(* IEC 61131-3 sources: plcassist-cli/packages/volt-lsp-iec/test-corpus/pro2193/Device/Plc Logic/Application/09 Misc/Library Manager/L_USPP_SignalProcessing, 27 files *)

(* ---- GETBOOLEANPROPERTY.fun ---- *)
FUNCTION GETBOOLEANPROPERTY : BOOL
VAR_INPUT
	STKEY : WSTRING;
END_VAR
END_FUNCTION

(* ---- GETCOMPANY.fun ---- *)
FUNCTION GETCOMPANY : WSTRING
END_FUNCTION

(* ---- GETNUMBERPROPERTY.fun ---- *)
FUNCTION GETNUMBERPROPERTY : DINT
VAR_INPUT
	STKEY : WSTRING;
END_VAR
END_FUNCTION

(* ---- GETTEXTPROPERTY.fun ---- *)
FUNCTION GETTEXTPROPERTY : WSTRING
VAR_INPUT
	STKEY : WSTRING;
END_VAR
END_FUNCTION

(* ---- GETTEXTPROPERTY2.fun ---- *)
FUNCTION GETTEXTPROPERTY2 : POINTER TO WSTRING
VAR_INPUT
	STKEY : WSTRING;
END_VAR
END_FUNCTION

(* ---- GETTITLE.fun ---- *)
FUNCTION GETTITLE : WSTRING
END_FUNCTION

(* ---- GETVERSION.fun ---- *)
FUNCTION GETVERSION : VERSION
END_FUNCTION

(* ---- GETVERSIONPROPERTY.fun ---- *)
FUNCTION GETVERSIONPROPERTY : VERSION
VAR_INPUT
	STKEY : WSTRING;
END_VAR
END_FUNCTION

(* ---- L_USPP_HLPPT1FILT.fun ---- *)
FUNCTION L_USPP_HLPPT1FILT : LREAL
VAR_INPUT
	LRVALUE : LREAL;
	LRINPUT : LREAL;
	LRNEW_N : LREAL;
END_VAR
END_FUNCTION

(* ---- GLOBALTEXTLIST.fb ---- *)
FUNCTION_BLOCK GLOBALTEXTLIST
VAR
	M_TEXTLISTFILE : STRING(255);
	_STNAMESPACE : STRING;
END_VAR
END_FUNCTION_BLOCK

(* ---- IMAGEPOOL.fb ---- *)
FUNCTION_BLOCK IMAGEPOOL
VAR
	M_STNAMESPACE : STRING(80);
	M_STHELPVARID : STRING;
	M_STHELPVARPATH : STRING(255);
	M_STHELP : STRING;
	M_REGISTERIMAGES : BOOL := TRUE;
END_VAR
END_FUNCTION_BLOCK

METHOD FB_INIT : BOOL
VAR_INPUT
	BINITRETAINS : BOOL;
	BINCOPYCODE : BOOL;
END_VAR
END_METHOD

METHOD FB_REINIT : BOOL
END_METHOD

METHOD FB_EXIT : BOOL
VAR_INPUT
	BINCOPYCODE : BOOL;
END_VAR
END_METHOD

(* ---- L_USPP_AVERAGEFILTER.fb ---- *)
FUNCTION_BLOCK L_USPP_AVERAGEFILTER EXTENDS L_USPP_Filter
VAR_INPUT
	LRFILTERTIME : LREAL;
	XCALCFILTERDELAY : BOOL := TRUE;
END_VAR
VAR_OUTPUT
	LRFILTERDELAY : LREAL;
END_VAR
VAR
	_ITFMEMORY : L_UBUP_IMemoryProvider;
	_DWDIM : DWORD;
	_DWBUFFERCOUNT : DWORD;
	_DWACTFILTERDEPTH : DWORD;
	_DWBUFFERSIZE : DWORD;
	_DWMEMSIZE : DWORD;
	_DWACTBUFFERPOS : DWORD;
	_DWPREVBUFFERPOS : DWORD;
	_DWVALIDDATA : DWORD;
	_ALRPTRBUFFER : ARRAY [0..(dwMaxDeriv + 1)] OF POINTER TO LREAL;
	_ONE_OVER_N : LREAL;
	_XFIRSTROUNDDONE : BOOL;
	_DWSTANDSTILLCNT : DWORD;
	_ALRFILTERED : ARRAY [0..dwMaxDeriv] OF LREAL;
END_VAR
END_FUNCTION_BLOCK

METHOD CYCLICACTION
VAR_INPUT
	ITFTIMINGCONTROLLER : L_UBUP.L_UBUP_ITimingController;
END_VAR
VAR_OUTPUT
	XCOMPLETE : BOOL;
	XABORT : BOOL;
	IERRORID : INT;
END_VAR
END_METHOD

METHOD RESETACTION
VAR_OUTPUT
	XCOMPLETE : BOOL;
END_VAR
END_METHOD

METHOD STARTACTION
VAR_OUTPUT
	XCOMPLETE : BOOL;
	IERRORID : INT;
END_VAR
END_METHOD

METHOD EVALMEMORYPROVIDER
VAR_INPUT
	ITFMEMORYPROVIDER : L_UBUP_IMemoryProvider;
END_VAR
END_METHOD

METHOD FB_INIT : BOOL
VAR_INPUT
	BINITRETAINS : BOOL;
	BINCOPYCODE : BOOL;
	DWDERIVS : DWORD;
	ITFMEMORY : L_UBUP_IMemoryProvider;
END_VAR
END_METHOD

METHOD FILTERDELAY : LREAL
VAR_INPUT
	LRROUNDS : LREAL;
	LRCYCLELENGTH : LREAL;
END_VAR
END_METHOD

METHOD DISTRIBUTEBUFFER
END_METHOD

METHOD FILTER
VAR_INPUT
	PLR : POINTER TO LREAL;
END_VAR
VAR_IN_OUT
	LRFILTERED : LREAL;
END_VAR
END_METHOD

METHOD FILTERDETECTOVERFLOW
VAR_INPUT
	LRNEXTPOS : LREAL;
	LRPREVPOS : LREAL;
	LRMODCYCLE : LREAL;
END_VAR
VAR_OUTPUT
	LRMODCYCLENEW : LREAL;
END_VAR
END_METHOD

METHOD FILTERMODULO
END_METHOD

METHOD FILTEROUTPUT
VAR_IN_OUT
	ALRFILTERED : ARRAY [0..dwMaxDeriv] OF LREAL;
	ALROUTPUT : ARRAY [0..dwMaxDeriv] OF LREAL;
END_VAR
END_METHOD

(* ---- L_USPP_AVERAGEFILTEREXPLICIT.fb ---- *)
FUNCTION_BLOCK L_USPP_AVERAGEFILTEREXPLICIT EXTENDS L_USPP_AverageFilter
END_FUNCTION_BLOCK

METHOD FB_INIT : BOOL
VAR_INPUT
	BINITRETAINS : BOOL;
	BINCOPYCODE : BOOL;
	DWDERIVS : DWORD;
	ITFMEMORY : L_UBUP_IMemoryProvider;
END_VAR
END_METHOD

METHOD FILTER
VAR_INPUT
	PLR : POINTER TO LREAL;
END_VAR
VAR_IN_OUT
	LRFILTERED : LREAL;
END_VAR
END_METHOD

METHOD FILTERMODULO
END_METHOD

(* ---- L_USPP_AVERAGEFILTERRECURSIVE.fb ---- *)
FUNCTION_BLOCK L_USPP_AVERAGEFILTERRECURSIVE EXTENDS L_USPP_AverageFilter
VAR
	_XALLOWMODULO : BOOL;
END_VAR
END_FUNCTION_BLOCK

METHOD STARTACTION
VAR_OUTPUT
	XCOMPLETE : BOOL;
	IERRORID : INT;
END_VAR
END_METHOD

METHOD FB_INIT : BOOL
VAR_INPUT
	BINITRETAINS : BOOL;
	BINCOPYCODE : BOOL;
	DWDERIVS : DWORD;
	ITFMEMORY : L_UBUP_IMemoryProvider;
	XALLOWMODULO : BOOL;
END_VAR
END_METHOD

METHOD FILTERROUNDSCOUNTING
END_METHOD

METHOD FILTER
VAR_INPUT
	PLR : POINTER TO LREAL;
END_VAR
VAR_IN_OUT
	LRFILTERED : LREAL;
END_VAR
END_METHOD

METHOD FILTERMODULO
END_METHOD

METHOD FILTEROUTPUT
VAR_IN_OUT
	ALRFILTERED : ARRAY [0..dwMaxDeriv] OF LREAL;
	ALROUTPUT : ARRAY [0..dwMaxDeriv] OF LREAL;
END_VAR
END_METHOD

(* ---- L_USPP_BUTTERWORTH2NDORDER.fb ---- *)
FUNCTION_BLOCK L_USPP_BUTTERWORTH2NDORDER
VAR_INPUT
	LRIN : LREAL;
	LRFILTERTIME : LREAL;
	LRSAMPLINGTIME : LREAL;
	XINITWITHFIRSTINPUTVALUE : BOOL;
END_VAR
VAR_OUTPUT
	LROUT : LREAL;
END_VAR
VAR
	_LRINITCYCLETIME : LREAL;
	_LRFILTERTIME : LREAL;
	LRTASKCYCLE : LREAL;
	LROMEGA : LREAL;
	ALRXINT : ARRAY [0..2] OF LREAL;
	ALRYINT : ARRAY [0..2] OF LREAL;
	LRB0 : LREAL;
	LRB1 : LREAL;
	LRB2 : LREAL;
	LRA0 : LREAL;
	LRA0INV : LREAL;
	LRA1 : LREAL;
	LRA2 : LREAL;
	LROMEGASQUARED : LREAL;
	C_LRSQRT2 : LREAL := SQRT(2);
END_VAR
END_FUNCTION_BLOCK

METHOD FB_INIT : BOOL
VAR_INPUT
	BINITRETAINS : BOOL;
	BINCOPYCODE : BOOL;
END_VAR
END_METHOD

(* ---- L_USPP_COMPARE.fb ---- *)
FUNCTION_BLOCK L_USPP_COMPARE
VAR_INPUT
	LRIN1 : LREAL := 0;
	LRIN2 : LREAL := 0;
	DWFUNCTION : DWORD := 0;
	LRTOLERANCE : LREAL := 0;
	LRHYSTERESIS : LREAL := 0;
END_VAR
VAR_OUTPUT
	XOUT : BOOL := FALSE;
	XERROR : BOOL := FALSE;
	EERRORID : L_IE1P_Error;
END_VAR
VAR
	LRINTHYSTERESIS : LREAL := 0;
	LRINTWINDOW : LREAL := 0;
	LRINTIN1 : LREAL := 0;
	LRINTIN2 : LREAL := 0;
	LRINTTEMP : LREAL := 0;
	OUTVAR : BOOL;
END_VAR
END_FUNCTION_BLOCK

(* ---- L_USPP_CURVE.fb ---- *)
FUNCTION_BLOCK L_USPP_CURVE
VAR_INPUT
	LRIN : LREAL;
	DWMODE : DWORD;
	ALRXVALUES : ARRAY [1..9] OF LREAL;
	ALRYVALUES : ARRAY [1..9] OF LREAL;
END_VAR
VAR_OUTPUT
	LROUT : LREAL;
	XERROR : BOOL := FALSE;
	EERRORID : L_IE1P_Error;
END_VAR
VAR
	DISTARTIDX : DINT;
	DIENDIDX : DINT;
	LRLASTIN : LREAL;
	LRINPUT : LREAL;
	DISTART : DINT;
	DIEND : DINT;
	DITMP32 : DINT;
	XNEGINPUT : BOOL;
	XSAVELASTIN : BOOL;
	TMP : LREAL;
	GETMAXCURVEPOINTS : INT := 9;
END_VAR
END_FUNCTION_BLOCK

METHOD GETVALIDDATA
END_METHOD

(* ---- L_USPP_DEADTIMEINT.fb ---- *)
FUNCTION_BLOCK L_USPP_DEADTIMEINT
VAR_INPUT
	XENABLE : BOOL;
	XOFFSETACTIVE : BOOL;
	LRDELAY : LREAL;
	LRCYCLETIME : LREAL;
	PBIN : POINTER TO BYTE;
	PBOUT : POINTER TO BYTE;
	DISIZEOFDATA : DINT;
END_VAR
VAR_OUTPUT
	XBUSY : BOOL;
	XBUFFERINITIALIZED : BOOL;
	XERROR : BOOL;
	EERRORID : L_IE1P_Error;
END_VAR
VAR
	_XENABLEOLD : BOOL;
	_XOFFSETACTIVE : BOOL;
	_UDISIZEINT : UDINT;
	_LRCYCLETIME : LREAL;
	_LRINITCYCLETIME : LREAL;
	_WBUFFERCNT_1 : WORD;
	_WBUFFERCNT_2 : WORD;
	_WBUFFERLENGTH : WORD;
	_LRDELAY : LREAL;
	_LRRES : LREAL;
	_WDELAY : WORD;
	_PTMP : POINTER TO BYTE;
	_ITFMEMPROVIDER : L_UBUP_IMemoryProvider;
	_PBBUFFER : POINTER TO BYTE;
	_UDIBUFFERSIZE : UDINT;
END_VAR
END_FUNCTION_BLOCK

METHOD FB_INIT : BOOL
VAR_INPUT
	BINITRETAINS : BOOL;
	BINCOPYCODE : BOOL;
	ITFMEMPROVIDER : L_UBUP_IMemoryProvider;
END_VAR
END_METHOD

METHOD EVALMEMORYPROVIDER
VAR_INPUT
	ITFMEMORYPROVIDER : L_UBUP_IMemoryProvider;
END_VAR
END_METHOD

(* ---- L_USPP_DELAY.fb ---- *)
FUNCTION_BLOCK L_USPP_DELAY
VAR_INPUT
	XIN : BOOL;
	DWFUNCTION : DWORD := 0;
	LRDELAYTIME : LREAL := 0.001;
END_VAR
VAR_OUTPUT
	XOUT : BOOL;
	XERROR : BOOL := FALSE;
	EERRORID : L_IE1P_Error;
END_VAR
VAR
	DWDELTICKS : DWORD;
	DWCOUNTER : DWORD;
	XINOLD : BOOL;
	DWTASKINTERVALL : DWORD;
	_LRINITCYCLETIME : LREAL;
END_VAR
END_FUNCTION_BLOCK

METHOD FB_INIT : BOOL
VAR_INPUT
	BINITRETAINS : BOOL;
	BINCOPYCODE : BOOL;
END_VAR
END_METHOD

(* ---- L_USPP_DIFFERENTIATE.fb ---- *)
FUNCTION_BLOCK L_USPP_DIFFERENTIATE
VAR_INPUT
	LRIN : LREAL;
	LRFILTERTIME : LREAL;
END_VAR
VAR_OUTPUT
	LROUT : LREAL;
END_VAR
VAR
	LRTASKCYCLE : LREAL;
	LRTEMP : LREAL;
	LRTIME : LREAL;
	LRINT : LREAL;
	_LRINITCYCLETIME : LREAL;
END_VAR
END_FUNCTION_BLOCK

METHOD FB_INIT : BOOL
VAR_INPUT
	BINITRETAINS : BOOL;
	BINCOPYCODE : BOOL;
END_VAR
END_METHOD

(* ---- L_USPP_FILTER.fb ---- *)
FUNCTION_BLOCK L_USPP_FILTER
VAR_INPUT
	XENABLE : BOOL;
	LRCYCLETIME : LREAL := L_UMTP_Math.L_UMTP_ValueIgnore;
	LRCYCLELENGTH : LREAL := L_UMTP_Math.L_UMTP_ValueIgnore;
	LRREFPOS : LREAL := L_UMTP_Math.L_UMTP_ValueIgnore;
	ALRIN : ARRAY [0..dwMaxDeriv] OF LREAL;
END_VAR
VAR_OUTPUT
	ALROUT : ARRAY [0..dwMaxDeriv] OF LREAL;
	XBUSY : BOOL;
	XERROR : BOOL;
	EERRORID : L_IE1P_Error;
END_VAR
VAR
	_LRCYCLELENGTH : LREAL;
	_LRCYCLELENGTHINV : LREAL;
	_LRCYCLETIME : LREAL;
	_XMODULO : BOOL;
	_MODEL : L_UBUP_BehaviourModel_LCon;
	DWMAXDERIV : DWORD := 3;
END_VAR
END_FUNCTION_BLOCK

METHOD REPLACE : L_IE1P_Error
VAR_INPUT
	ACTFILTER : REFERENCE TO L_USPP_Filter;
END_VAR
END_METHOD

METHOD CYCLICACTION
VAR_INPUT
	ITFTIMINGCONTROLLER : L_UBUP.L_UBUP_ITimingController;
END_VAR
VAR_OUTPUT
	XCOMPLETE : BOOL;
	XABORT : BOOL;
	IERRORID : INT;
END_VAR
END_METHOD

METHOD FINALIZEACTION
VAR_INPUT
	XABORTPROPOSED : BOOL;
	IERRORIDPROPOSED : INT;
END_VAR
VAR_OUTPUT
	XCOMPLETE : BOOL;
	XABORT : BOOL;
	IERRORID : INT;
END_VAR
END_METHOD

METHOD RESETACTION
VAR_OUTPUT
	XCOMPLETE : BOOL;
END_VAR
END_METHOD

METHOD STARTACTION
VAR_OUTPUT
	XCOMPLETE : BOOL;
	IERRORID : INT;
END_VAR
END_METHOD

(* ---- L_USPP_INTEGRATE.fb ---- *)
FUNCTION_BLOCK L_USPP_INTEGRATE
VAR_INPUT
	LRIN : LREAL;
	XLOADSTARTVALUE : BOOL;
	LRSTARTVALUE : LREAL;
END_VAR
VAR_OUTPUT
	LROUT : LREAL;
END_VAR
VAR
	LRTASKCYCLE : LREAL;
	LRTEMP : LREAL;
	_LRINITCYCLETIME : LREAL;
END_VAR
END_FUNCTION_BLOCK

METHOD FB_INIT : BOOL
VAR_INPUT
	BINITRETAINS : BOOL;
	BINCOPYCODE : BOOL;
END_VAR
END_METHOD

(* ---- L_USPP_OSCILLATOR.fb ---- *)
FUNCTION_BLOCK L_USPP_OSCILLATOR
VAR_INPUT
	XENABLE : BOOL;
	LRTIMEHIGH : LREAL := 0.001;
	LRTIMELOW : LREAL := 0.001;
END_VAR
VAR_OUTPUT
	XOUT : BOOL;
END_VAR
VAR
	DWTASKINTERVAL : DWORD;
	DWTIMEHIGH : DWORD;
	DWTIMELOW : DWORD;
	DWTIMEPERIOD : DWORD;
	DWCOUNTER : DWORD;
	_LRINITCYCLETIME : LREAL;
END_VAR
END_FUNCTION_BLOCK

METHOD FB_INIT : BOOL
VAR_INPUT
	BINITRETAINS : BOOL;
	BINCOPYCODE : BOOL;
END_VAR
END_METHOD

(* ---- L_USPP_PIDREGLER.fb ---- *)
FUNCTION_BLOCK L_USPP_PIDREGLER EXTENDS L_USPP_Filter
END_FUNCTION_BLOCK

METHOD FB_INIT : BOOL
VAR_INPUT
	BINITRETAINS : BOOL;
	BINCOPYCODE : BOOL;
END_VAR
END_METHOD

METHOD CYCLICACTION
VAR_INPUT
	ITFTIMINGCONTROLLER : L_UBUP.L_UBUP_ITimingController;
END_VAR
VAR_OUTPUT
	XCOMPLETE : BOOL;
	XABORT : BOOL;
	IERRORID : INT;
END_VAR
END_METHOD

(* ---- L_USPP_PT1FILTER.fb ---- *)
FUNCTION_BLOCK L_USPP_PT1FILTER
VAR_INPUT
	LRIN : LREAL;
	LRDELAYTIME : LREAL := 0.0;
END_VAR
VAR_OUTPUT
	LROUT : LREAL;
	XERROR : BOOL := FALSE;
	EERRORID : L_IE1P_Error;
END_VAR
VAR
	LRTIME : LREAL;
	LRTASKCYCLE : LREAL;
	LRTEMP : LREAL;
	_LRINITCYCLETIME : LREAL;
END_VAR
END_FUNCTION_BLOCK

METHOD FB_INIT : BOOL
VAR_INPUT
	BINITRETAINS : BOOL;
	BINCOPYCODE : BOOL;
END_VAR
END_METHOD

(* ---- L_USPP_PT2FILTER.fb ---- *)
FUNCTION_BLOCK L_USPP_PT2FILTER EXTENDS L_USPP_Filter
VAR_INPUT
	LRT1 : LREAL;
	LRT2 : LREAL;
	LRV : LREAL;
END_VAR
VAR
	_LRA : LREAL;
	_LRB : LREAL;
	_LRK : LREAL;
	_LRT : LREAL;
	_LRT1 : LREAL;
	_LRT2 : LREAL;
END_VAR
END_FUNCTION_BLOCK

METHOD CYCLICACTION
VAR_INPUT
	ITFTIMINGCONTROLLER : L_UBUP.L_UBUP_ITimingController;
END_VAR
VAR_OUTPUT
	XCOMPLETE : BOOL;
	XABORT : BOOL;
	IERRORID : INT;
END_VAR
END_METHOD

METHOD STARTACTION
VAR_OUTPUT
	XCOMPLETE : BOOL;
	IERRORID : INT;
END_VAR
END_METHOD

(* ---- L_USPP_SELECT.fb ---- *)
FUNCTION_BLOCK L_USPP_SELECT
VAR_INPUT
	LRIN1 : LREAL := 0;
	LRIN2 : LREAL := 0;
	XSELECTIN2 : BOOL := FALSE;
END_VAR
VAR_OUTPUT
	LROUT : LREAL := 0;
END_VAR
END_FUNCTION_BLOCK
